Fanuc KAREL source: ka00089.KL

-- PROVISIONAL review KL for V770-1; original PC SHA256 81755dd3d1747a1d2fb14a5ab59caa85c5e6d280c415bd5551d7be8b9c5c41b0
-- Incomplete behavior may be omitted. Consult companion uncertainty JSON. Do not deploy.
PROGRAM KA00089
%NOLOCKGROUP
-- UNRESOLVED_DECL SRC type=000199
-- UNRESOLVED_DECL DST type=000101
BEGIN
  -- UNRESOLVED_PC offsets 5-25; opcodes 49,7E,4A
  -- UNRESOLVED_PC offsets 30-34; opcodes 7F
END KA00089
